(* IEC 61131-3 sources: codesys-to-astra/src/POUs/F_C2aMx210Status, 2 files *)

(* ---- F_C2aMx210Status.decl.st ---- *)
// Назначение: код ошибки датчика МВ210-101 (РЭ v1.41, табл. 6.9, с. 36) -> E_C2aMx210Status; код вне
//             таблицы — Ok (передаётся результат измерения).
// Автор:      kr0nsch
// Версия:     0.1.0
// Документ:   docs/IO.md
FUNCTION F_C2aMx210Status : E_C2aMx210Status
VAR_INPUT
    bCode : BYTE;      // код из регистра значения
END_VAR

(* ---- F_C2aMx210Status.impl.st ---- *)
CASE bCode OF
    16#F0: F_C2aMx210Status := E_C2aMx210Status.Invalid;
    16#F6: F_C2aMx210Status := E_C2aMx210Status.NotReady;
    16#F7: F_C2aMx210Status := E_C2aMx210Status.SensorOff;
    16#F8: F_C2aMx210Status := E_C2aMx210Status.ColdJunctionHigh;
    16#F9: F_C2aMx210Status := E_C2aMx210Status.ColdJunctionLow;
    16#FA: F_C2aMx210Status := E_C2aMx210Status.TooHigh;
    16#FB: F_C2aMx210Status := E_C2aMx210Status.TooLow;
    16#FC: F_C2aMx210Status := E_C2aMx210Status.ShortCircuit;
    16#FD: F_C2aMx210Status := E_C2aMx210Status.SensorBreak;
    16#FE: F_C2aMx210Status := E_C2aMx210Status.AdcFailure;
    16#FF: F_C2aMx210Status := E_C2aMx210Status.BadCalibration;
ELSE
    F_C2aMx210Status := E_C2aMx210Status.Ok;
END_CASE
